FUNCTION FC 1 : VOID
BEGIN
NETWORK
      U I 0.0
END_FUNCTION
